// TIA Portal V20 export
Screen "Pop-up_PRODDATA_LV_LEGEND_Popup"  340x273
  ScreenItem "Background" at 0,0 size 340x273  Type=HmiRectangle
  ScreenItem "Textfeld_Legende" at 1,1 size 328x25  Type=HmiTextBox
  ScreenItem "Textfeld_11" at 70,178 size 255x89  Type=HmiTextBox
  ScreenItem "Textfeld_8" at 10,226 size 55x30  Type=HmiTextBox
  ScreenItem "Textfeld_9" at 23,207 size 30x20  Type=HmiTextBox
  ScreenItem "Textfeld_13" at 10,178 size 55x30  Type=HmiTextBox
  ScreenItem "Textfeld_12" at 10,38 size 208x25  Type=HmiTextBox
  ScreenItem "Textfeld_15" at 10,63 size 315x40  Type=HmiTextBox
  ScreenItem "Textfeld_5" at 10,105 size 55x30  Type=HmiTextBox
  ScreenItem "Textfeld_6" at 70,101 size 268x71  Type=HmiTextBox
  ScreenItem "Textfeld_7" at 10,138 size 55x30  Type=HmiTextBox
  ScreenItem "Cancel Mode" at 249,1 size 90x60  Type=HmiButton
